SUBAPPLICATION Uebung_162_AX (* Übung zu DS18B20: Temperatur messen, Q1 über 25 °C *)
  (* Standard: 61499-2; Description: Copyright (c) 2026 Meisterschulen am Ostbahnhof This program and the accompanying materials are made available under the terms of the Eclipse Public License 2.0 which is available at https://www.eclipse.org/legal/epl-2.0/ SPDX-License-Identifier: EPL-2.0 *)
  (* Version 1.0, 2026-11-26, Franz Höpfinger, Meisterschulen am Ostbahnhof, initial API and implementation and/or initial documentation *)
  PACKAGE Uebungen;
  IMPORT logiBUS::io::DQ::logiBUS_DO::Output_Q1;
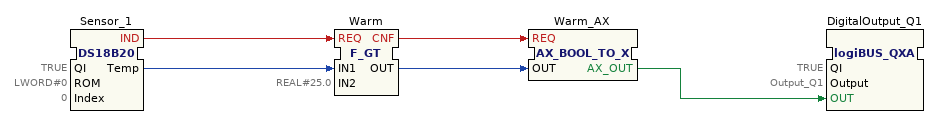
  (* Temperatursensor DS18B20 (logiBUS_onewire) am Trainer20: Datenleitung GPIO3, externer Pull-up 4,7 kOhm empfohlen. IND nach jeder Messrunde (ca. 1 s, 12 Bit). Q1 an = wärmer als 25 °C (Sensor in der Hand anwärmen). Watch: Temp (°C), QO (TRUE = Temp gültig), STATUS, ROMO (ROM-Code des Sensors, für Übung 162b notieren). STATUS z. B. 'sensor not found', 'power-on value 85 C' (erste Messung noch nicht fertig), 'no 1-Wire bus on this board'. Weiter: Übung 162b (zwei Sensoren, einer per ROM-Code festgehalten). *)
  FBS
    Sensor_1 : logiBUS::onewire::DS18B20(QI := TRUE, ROM := LWORD#0, Index := 0); (* erster Sensor am Bus (Index 0) *)
    Warm : iec61131::comparison::F_GT(IN2 := REAL#25.0); (* Temp über 25 °C? *)
    Warm_AX : adapter::conversion::unidirectional::AX_BOOL_TO_X;
    DigitalOutput_Q1 : logiBUS::io::DQ::logiBUS_QXA(QI := TRUE, Output := Output_Q1); (* an = wärmer als 25 °C *)
  END_FBS
  EVENT_CONNECTIONS
    Sensor_1.IND TO Warm.REQ;
    Warm.CNF TO Warm_AX.REQ;
  END_CONNECTIONS
  DATA_CONNECTIONS
    Sensor_1.Temp TO Warm.IN1;
    Warm.OUT TO Warm_AX.OUT;
  END_CONNECTIONS
  ADAPTER_CONNECTIONS
    Warm_AX.AX_OUT TO DigitalOutput_Q1.OUT;
  END_CONNECTIONS
END_SUBAPPLICATION
